Fanuc KAREL source: KC00058.KL

PROGRAM KC00058
%NOLOCKGROUP
%ENVIRONMENT DEBUG
VAR
  I: INTEGER
  J: INTEGER
  K: INTEGER
  R: REAL
  B: BOOLEAN
  S: STRING[80]
  T: STRING[80]
  P: PATH
  Q: PATH
  AI: ARRAY[8] OF INTEGER
  AB: ARRAY[244] OF BYTE
BEGIN
  CHECK_STACK(B,B,I)
END KC00058
